// TIA Portal V19 export
// export: Created 2026-10-15T09:44:24.2356284Z, ExportSetting WithDefaults, DisplayName Totally Integrated Automation Portal, DisplayVersion V19, DisplayName TIA Portal Openness, DisplayVersion V19, DisplayName TIA Portal Version Control Interface, DisplayVersion V19, DisplayName STEP 7 Professional, DisplayVersion V19, DisplayName STEP 7 Safety, DisplayVersion V19, DisplayName WinCC Basic/Comfort/Advanced, DisplayVersion V19, DisplayName WinCC Unified, DisplayVersion V19
FUNCTION "ROLL_PB14" : Void   // FC22, SCL
{ S7_Optimized_Access := 'TRUE' }
VERSION : 0.1
// stored: AutoNumber true, IsIECCheckEnabled false, SetENOAutomatically false, UDAEnableTagReadback false
   VAR_TEMP
      r : Bool;
      a1 : Word;
      a2 : Word;
      activeDataBlock : Int;
      comparisonResults : Array[0..0] of Bool;
   END_VAR
BEGIN

   #r := FALSE;
   #a1 := W#16#0000;
   #a2 := W#16#0000;
   #activeDataBlock := 0;
   // PB14, STEP 5 network 1
   #activeDataBlock := 15;
   // PB14, STEP 5 network 2
   #r := ((NOT "ROLL_State".M[37, 5]) AND (NOT "ROLL_State".M[53, 2]) AND (NOT "ROLL_State".M[53, 3]) AND (((NOT "ROLL_State".S5Timers[21].Q) AND "ROLL_IO".Input[123, 4] AND "ROLL_State".M[31, 4]) OR ("ROLL_State".M[70, 4] AND "ROLL_State".S5Timers[45].Q) OR "ROLL_State".M[37, 7] OR "ROLL_State".M[53, 4] OR "ROLL_State".M[70, 7]) AND ((NOT "ROLL_State".S5Timers[95].Q) OR "ROLL_State".M[53, 4]) AND "ROLL_State".M[31, 5] AND "ROLL_State".M[35, 2]);
   "ROLL_State".M[64, 0] := #r;
   // PB14, STEP 5 network 3
   #r := (((NOT "ROLL_State".M[31, 4]) AND (NOT "ROLL_State".M[31, 5]) AND "ROLL_IO".Input[125, 4]) OR ((((NOT "ROLL_IO".Output[113, 4]) AND "ROLL_IO".Output[113, 5] AND "ROLL_State".M[72, 1]) OR "ROLL_State".M[53, 4]) AND "ROLL_State".M[31, 5] AND "ROLL_State".M[35, 2]));
   "ROLL_State".M[64, 1] := #r;
   // PB14, STEP 5 network 4
   #r := ("ROLL_IO".Input[123, 4] AND "ROLL_State".S5Timers[20].Q);
   IF #r THEN
       "ROLL_State".M[64, 4] := TRUE;
   END_IF;
   #r := (((NOT "ROLL_IO".Output[113, 3]) AND (NOT "ROLL_IO".Input[123, 4])) OR (NOT "ROLL_State".M[31, 5]));
   IF #r THEN
       "ROLL_State".M[64, 4] := FALSE;
   END_IF;
   // PB14, STEP 5 network 5
   #r := "ROLL_State".M[37, 5];
   IF #r THEN
       "ROLL_State".M[64, 5] := TRUE;
   END_IF;
   #r := ((NOT "ROLL_State".M[31, 5]) OR "ROLL_State".M[39, 5]);
   IF #r THEN
       "ROLL_State".M[64, 5] := FALSE;
   END_IF;
   // PB14, STEP 5 network 6
   #r := ((("ROLL_State".M[40, 2] OR "ROLL_State".M[44, 7] OR "ROLL_State".M[50, 6]) AND "ROLL_State".M[63, 1]) OR "ROLL_State".M[41, 6] OR "ROLL_State".M[43, 2] OR "ROLL_State".M[44, 7] OR "ROLL_State".M[46, 2] OR "ROLL_State".M[47, 6] OR "ROLL_State".M[49, 2]);
   "ROLL_State".M[65, 0] := #r;
   // PB14, STEP 5 network 7
   #r := ("ROLL_IO".Input[12, 5] AND "ROLL_IO".Input[12, 7] AND "ROLL_State".M[52, 0] AND "ROLL_State".M[63, 1]);
   "ROLL_State".M[65, 5] := #r;
   // PB14, STEP 5 network 8
   #r := (((NOT "ROLL_IO".Input[11, 0]) AND "ROLL_State".M[52, 0]) OR ((NOT "ROLL_IO".Input[11, 1]) AND "ROLL_State".M[40, 2]) OR ((NOT "ROLL_IO".Input[11, 2]) AND "ROLL_State".M[41, 6]) OR ((NOT "ROLL_IO".Input[11, 3]) AND "ROLL_State".M[43, 2]) OR ((NOT "ROLL_IO".Input[11, 4]) AND "ROLL_State".M[44, 7]) OR ((NOT "ROLL_IO".Input[119, 6]) AND "ROLL_State".M[46, 2]) OR ((NOT "ROLL_IO".Input[119, 7]) AND "ROLL_State".M[47, 6]) OR ((NOT "ROLL_IO".Input[120, 0]) AND "ROLL_State".M[49, 2]) OR ((NOT "ROLL_IO".Input[120, 1]) AND "ROLL_State".M[50, 6]));
   "ROLL_State".M[65, 6] := #r;
   // PB14, STEP 5 network 9
   #r := (("ROLL_IO".Input[11, 0] AND "ROLL_State".M[40, 0]) OR ("ROLL_IO".Input[11, 1] AND "ROLL_State".M[41, 0]) OR ("ROLL_IO".Input[11, 2] AND "ROLL_State".M[42, 4]) OR ("ROLL_IO".Input[11, 3] AND "ROLL_State".M[44, 0]) OR ("ROLL_IO".Input[11, 4] AND "ROLL_State".M[45, 5]) OR ("ROLL_IO".Input[119, 6] AND "ROLL_State".M[47, 0]) OR ("ROLL_IO".Input[119, 7] AND "ROLL_State".M[48, 4]) OR ("ROLL_IO".Input[120, 0] AND "ROLL_State".M[50, 0]) OR ("ROLL_IO".Input[120, 1] AND "ROLL_State".M[51, 3]));
   "ROLL_State".M[66, 2] := #r;
   // PB14, STEP 5 network 10
   #r := (("ROLL_State".M[66, 2] OR "ROLL_State".M[68, 2]) AND "ROLL_IO".Input[11, 6]);
   "ROLL_State".M[66, 4] := #r;
   // PB14, STEP 5 network 11
   #r := (("ROLL_IO".Input[11, 1] AND "ROLL_State".M[40, 4]) OR ("ROLL_IO".Input[11, 2] AND "ROLL_State".M[42, 0]) OR ("ROLL_IO".Input[11, 3] AND "ROLL_State".M[43, 4]) OR ("ROLL_IO".Input[11, 4] AND "ROLL_State".M[45, 1]) OR ("ROLL_IO".Input[119, 6] AND "ROLL_State".M[46, 4]) OR ("ROLL_IO".Input[119, 7] AND "ROLL_State".M[48, 0]) OR ("ROLL_IO".Input[120, 0] AND "ROLL_State".M[49, 4]) OR ("ROLL_IO".Input[120, 1] AND "ROLL_State".M[51, 0]));
   "ROLL_State".M[66, 5] := #r;
   // PB14, STEP 5 network 12
   #r := (((NOT "ROLL_IO".Input[12, 1]) OR (NOT "ROLL_IO".Input[12, 7])) AND "ROLL_IO".Input[11, 0] AND "ROLL_State".M[52, 2]);
   "ROLL_State".M[66, 6] := #r;
   // PB14, STEP 5 network 13
   #r := (("ROLL_State".M[66, 5] OR "ROLL_State".M[66, 6] OR "ROLL_State".M[68, 3]) AND "ROLL_IO".Input[11, 6]);
   "ROLL_State".M[66, 7] := #r;
   // PB14, STEP 5 network 14
   #r := ((NOT "ROLL_IO".Output[113, 3]) AND (NOT "ROLL_State".M[9, 3]) AND "ROLL_IO".Input[124, 5] AND "ROLL_State".M[39, 6]);
   "ROLL_State".M[67, 0] := #r;
   // PB14, STEP 5 network 15
   #r := ((NOT "ROLL_IO".Output[113, 3]) AND (NOT "ROLL_State".M[9, 3]) AND "ROLL_IO".Input[124, 5] AND "ROLL_State".M[53, 0]);
   "ROLL_State".M[67, 1] := #r;
   // PB14, STEP 5 network 16
   #r := ((NOT "ROLL_IO".Input[124, 5]) AND "ROLL_IO".Input[124, 1] AND "ROLL_State".M[39, 4]);
   "ROLL_State".M[67, 5] := #r;
   // PB14, STEP 5 network 17
   #r := ((NOT "ROLL_IO".Input[124, 4]) AND "ROLL_IO".Input[124, 1] AND "ROLL_State".M[53, 2]);
   "ROLL_State".M[67, 6] := #r;
   // PB14, STEP 5 network 18
   #r := ((("ROLL_IO".Input[5, 1] AND "ROLL_State".M[40, 5]) OR ("ROLL_State".M[0, 3] AND "ROLL_State".M[45, 2]) OR "ROLL_State".M[42, 1] OR "ROLL_State".M[43, 5] OR "ROLL_State".M[46, 5] OR "ROLL_State".M[48, 1] OR "ROLL_State".M[49, 5]) AND "ROLL_State".M[111, 3]);
   "ROLL_State".M[68, 0] := #r;
   // PB14, STEP 5 network 19
   #r := ((NOT "ROLL_State".S5Timers[25].Q) AND (("ROLL_IO".Input[12, 1] AND "ROLL_IO".Input[12, 7]) OR "ROLL_State".M[68, 2]) AND ("ROLL_State".M[68, 2] OR "ROLL_State".S5Timers[24].Q) AND "ROLL_State".M[68, 0]);
   "ROLL_State".M[68, 2] := #r;
   // PB14, STEP 5 network 20
   #r := (((NOT "ROLL_IO".Input[12, 1]) OR (NOT "ROLL_IO".Input[12, 7])) AND ("ROLL_State".M[68, 3] OR "ROLL_State".S5Timers[24].Q) AND "ROLL_State".M[68, 0]);
   "ROLL_State".M[68, 3] := #r;
   // PB14, STEP 5 network 21
   #a2 := #a1;
   #a1 := "ROLL_GetDW"(DbNumber := #activeDataBlock, Index := 24);
   #r := ((NOT "ROLL_State".M[68, 2]) AND (NOT "ROLL_State".M[68, 3]));
   "ROLL_TimerOp"(Number := 24,
                  Operation := 0,
                  Signal := #r,
                  Preset := #a1);
   // PB14, STEP 5 network 22
   #a2 := #a1;
   #a1 := "ROLL_GetDW"(DbNumber := #activeDataBlock, Index := 25);
   #r := "ROLL_State".M[68, 2];
   "ROLL_TimerOp"(Number := 25,
                  Operation := 0,
                  Signal := #r,
                  Preset := #a1);
   // PB14, STEP 5 network 23
   RETURN;
END_FUNCTION
